METHOD Work : E_PROGRESS // commands TransportUnit to TRANSPORT_START
VAR_INPUT
  Execute     : BOOL;
END_VAR
VAR_INST
  _nErrorId   : UDINT;
  _eState     : E_PROGRESS;
END_VAR
//-----------------------------------------------------------------------------
IF NOT Execute 
THEN 
	_eState                       := E_PROGRESS.PROGRESS_INIT; 
END_IF 
//-----------------------------------------------------------------------------
IF NOT Check() 
THEN 
	Work                          := E_PROGRESS.PROGRESS_ERROR; 
	RETURN; 
END_IF
//-----------------------------------------------------------------------------
//-----------------------------------------------------------------------------
CASE _eState
OF
  E_PROGRESS.PROGRESS_INIT:
    IF Execute
    THEN
      _nErrorId                 := 0;

      _XtsTransportCtrl.Cmd     := E_XTS_TRANSPORT_CTRL.CMD_NULL;
      _eState                   := E_PROGRESS.PROGRESS_BUSY;

      IF (_MessageLevel > E_MessageType.eMessageError)
      THEN
        _stMsg.eType            := E_MessageType.eMessageInfo;
        _stMsg.eSubdevice       := e_Subdevice.Application_Work;
        _stMsg.iErrorNumber     := 0;
        _stMsg.sText            := concat(TO_STRING(_eState), ': ');
        f_MessageSet(_stMsg);
      END_IF
    END_IF
  //-----------------------------------------------------------------------------
  //-----------------------------------------------------------------------------
  E_PROGRESS.PROGRESS_BUSY:
    _XtsTransportCtrl.Cmd       := E_XTS_TRANSPORT_CTRL.CMD_TRANSPORT_START;

    IF (_XtsTransportState.State = E_XTS_TRANSPORT_STATE.TRANSPORT_START + E_PROGRESS.PROGRESS_ERROR)
    THEN
      _eState                   := E_PROGRESS.PROGRESS_ERROR;
      _nErrorId                 := _XtsTransportState.GroupInfo.GroupErrorId; 

    ELSIF (_XtsTransportState.State = E_XTS_TRANSPORT_STATE.TRANSPORT_START + E_PROGRESS.PROGRESS_DONE)
    THEN
      _eState                   := E_PROGRESS.PROGRESS_PREPARE;
    END_IF
  //-----------------------------------------------------------------------------
  // spare states: 
  //  - the work is done for the YardMaster
  //  - you can now work on the CTRL/STATE structures of the Instances
  //-----------------------------------------------------------------------------
  E_PROGRESS.PROGRESS_PREPARE:
    _eState                     := E_PROGRESS.PROGRESS_STARTUP;
  //---------------------------------------------------------------------------------------------------------------
  //---------------------------------------------------------------------------------------------------------------
  E_PROGRESS.PROGRESS_STARTUP:
    _eState                     := E_PROGRESS.PROGRESS_CHECK;
  //---------------------------------------------------------------------------------------------------------------
  //---------------------------------------------------------------------------------------------------------------
  E_PROGRESS.PROGRESS_CHECK:
    _eState                     := E_PROGRESS.PROGRESS_OCCUPIED;
  //---------------------------------------------------------------------------------------------------------------
  //---------------------------------------------------------------------------------------------------------------
  E_PROGRESS.PROGRESS_OCCUPIED:
    _eState                     := E_PROGRESS.PROGRESS_WORKING;
  //---------------------------------------------------------------------------------------------------------------
  //---------------------------------------------------------------------------------------------------------------
  E_PROGRESS.PROGRESS_WORKING:
    _eState                     := E_PROGRESS.PROGRESS_STILL_WORKING;
  //---------------------------------------------------------------------------------------------------------------
  //---------------------------------------------------------------------------------------------------------------
  E_PROGRESS.PROGRESS_STILL_WORKING:
    _eState                     := E_PROGRESS.PROGRESS_DONE;

    IF (_MessageLevel > E_MessageType.eMessageError)
    THEN
      _stMsg.eType              := E_MessageType.eMessageInfo;
      _stMsg.eSubdevice         := e_Subdevice.Application_Work;
      _stMsg.iErrorNumber       := 0;
      _stMsg.sText              := concat(TO_STRING(_eState), ': ');
      f_MessageSet(_stMsg);
    END_IF

END_CASE
//-----------------------------------------------------------------------------
//-----------------------------------------------------------------------------

Work                            := _eState;
END_METHOD

PROPERTY XtsTransportCtrl : REFERENCE TO ST_XTS_TRANSPORT_CTRL
SET
_XtsTransportCtrl REF= XtsTransportCtrl;
END_SET
END_PROPERTY

PROPERTY XtsTransportState : REFERENCE TO ST_XTS_TRANSPORT_STATE
SET
_XtsTransportState REF= XtsTransportState;
END_SET
END_PROPERTY

END_FUNCTION_BLOCK

// ---- _MSG/f_MessageSet.TcPOU
FUNCTION f_MessageSet : BOOL
VAR_INPUT
  stMessage     : ST_Message;
END_VAR
VAR
  _uiIndex      : UINT;
  _MainDevice   : e_Device;
  _nModRes      : UDINT;     // residual after modulo
END_VAR

stMessage.tTime                     := GVL_MSG_XTS.sLocalTime;

// why here? so all calls to this function may stay the same
_nModRes                            := stMessage.eDevice MOD e_Device.General;
_MainDevice                         := stMessage.eDevice - _nModRes;

CASE _MainDevice
OF
  //--------------------------------------------------------------------------------
  e_device.DataProduct:
    // this is your data, if you choose to use this message system
    FOR _uiIndex := 1 TO GVL_MSG_XTS.MAX_MESSAGE
    DO
      IF (GVL_MSG_XTS.ProductMessages[_uiIndex].eType = e_MessageType.eMessageEmpty)
      THEN
        GVL_MSG_XTS.ProductMessages[_uiIndex]      := stMessage;
        GVL_MSG_XTS.MessageProductIndex            := _uiIndex;
        EXIT;
      END_IF
    END_FOR
  
    IF (stMessage.eType = E_MessageType.eMessageError)
    THEN
      // in case of error: increment counter
      GVL_MSG_XTS.MessageProductError              := GVL_MSG_XTS.MessageProductError + 1;
    END_IF
  //--------------------------------------------------------------------------------
  e_Device.Process,
  e_Device.Application:
    FOR _uiIndex := 1 TO GVL_MSG_XTS.MAX_MESSAGE
    DO
      IF (GVL_MSG_XTS.ApplicationMessages[_uiIndex].eType = e_MessageType.eMessageEmpty)
      THEN
        GVL_MSG_XTS.ApplicationMessages[_uiIndex]  := stMessage;    // yes, we grab global values directly, only here
        GVL_MSG_XTS.MessageApplicationIndex        := _uiIndex;
        EXIT;
      END_IF
    END_FOR
    IF (stMessage.eType = E_MessageType.eMessageError)
    THEN
      // in case of error: increment counter
      GVL_MSG_XTS.MessageApplicationError          := GVL_MSG_XTS.MessageApplicationError + 1;
    END_IF
  //--------------------------------------------------------------------------------
  e_Device.MetricsXts:
    FOR _uiIndex := 1 TO GVL_MSG_XTS.MAX_MESSAGE
    DO
      IF (GVL_MSG_XTS.MetricsMessages[_uiIndex].eType = e_MessageType.eMessageEmpty)
      THEN
        GVL_MSG_XTS.MetricsMessages[_uiIndex]      := stMessage;    // yes, we grab global values directly, only here
        GVL_MSG_XTS.MessageMetricsIndex            := _uiIndex;
        EXIT;
      END_IF
    END_FOR
    IF (stMessage.eType = E_MessageType.eMessageError)
    THEN
      // in case of error: increment counter
      GVL_MSG_XTS.MessageMetricsError              := GVL_MSG_XTS.MessageMetricsError + 1;
    END_IF
  //--------------------------------------------------------------------------------
  e_Device.MetricsAxis:
    FOR _uiIndex := 1 TO GVL_MSG_XTS.MAX_MESSAGE
    DO
      IF (GVL_MSG_AXIS.MetricMessages[_uiIndex].eType = e_MessageType.eMessageEmpty)
      THEN
        GVL_MSG_AXIS.MetricMessages[_uiIndex]  := stMessage;    // yes, we grab global values directly, only here
        GVL_MSG_AXIS.MessageMetricIndex        := _uiIndex;
        EXIT;
      END_IF
    END_FOR
    IF (stMessage.eType = E_MessageType.eMessageError)
    THEN
      // in case of error: increment counter
      GVL_MSG_AXIS.MessageMetricError          := GVL_MSG_AXIS.MessageMetricError + 1;
    END_IF
  //--------------------------------------------------------------------------------
  e_Device.Axis,
  e_Device.XfcAxis,
  e_device.XfcTouchProbe,
  e_device.XfcTriggerBox,
  e_Device.Camming,
  e_device.NciChannel,
  e_device.NciChannelCtrl:
    FOR _uiIndex := 1 TO GVL_MSG_XTS.MAX_MESSAGE
    DO
      IF (GVL_MSG_AXIS.MotionMessages[_uiIndex].eType = e_MessageType.eMessageEmpty)
      THEN
        GVL_MSG_AXIS.MotionMessages[_uiIndex]  := stMessage;    // yes, we grab global values directly, only here
        GVL_MSG_AXIS.MessageMotionIndex        := _uiIndex;
        EXIT;
      END_IF
    END_FOR
    IF (stMessage.eType = E_MessageType.eMessageError)
    THEN
      // in case of error: increment counter
      GVL_MSG_AXIS.MessageMotionError           := GVL_MSG_AXIS.MessageMotionError + 1;
    END_IF
  //--------------------------------------------------------------------------------
ELSE
  CASE stMessage.eDevice
  OF
    Device_MainApplication,
    Device_XmlData,              
    Device_Utilities:
      FOR _uiIndex := 1 TO GVL_MSG_XTS.MAX_MESSAGE
      DO
        IF (GVL_MSG_XTS.ApplicationMessages[_uiIndex].eType = e_MessageType.eMessageEmpty)
        THEN
          GVL_MSG_XTS.ApplicationMessages[_uiIndex]:= stMessage;    // yes, we grab global values directly, only here
          GVL_MSG_XTS.MessageApplicationIndex      := _uiIndex;
          EXIT;
        END_IF
      END_FOR
      IF (stMessage.eType = E_MessageType.eMessageError)
      THEN
        // in case of error: increment counter
        GVL_MSG_XTS.MessageApplicationError        := GVL_MSG_XTS.MessageApplicationError + 1;
      END_IF

    Device_MainAxis,
    Device_Nci,
    Device_Cam,
    Device_Functions,
    Device_FlyingSaw,
    Device_ParameterSelector:     // PLC_MOTION
      FOR _uiIndex := 1 TO GVL_MSG_XTS.MAX_MESSAGE
      DO
        IF (GVL_MSG_AXIS.MotionMessages[_uiIndex].eType = e_MessageType.eMessageEmpty)
        THEN
          GVL_MSG_AXIS.MotionMessages[_uiIndex]:= stMessage;    // yes, we grab global values directly, only here
          GVL_MSG_AXIS.MessageMotionIndex      := _uiIndex;
          EXIT;
        END_IF
      END_FOR
      IF (stMessage.eType = E_MessageType.eMessageError)
      THEN
        // in case of error: increment counter
        GVL_MSG_AXIS.MessageMotionError        := GVL_MSG_AXIS.MessageMotionError + 1;
      END_IF

    Device_Main,
    Device_MoverSelector:
      FOR _uiIndex := 1 TO GVL_MSG_XTS.MAX_MESSAGE
      DO
        IF (GVL_MSG_XTS.TransportMessages[_uiIndex].eType = e_MessageType.eMessageEmpty)
        THEN
          GVL_MSG_XTS.TransportMessages[_uiIndex]  := stMessage;
          GVL_MSG_XTS.MessageTransportIndex        := _uiIndex;
          EXIT;
        END_IF
      END_FOR
  ELSE    
    //--------------------------------------------------------------------------------
    FOR _uiIndex := 1 TO GVL_MSG_XTS.MAX_MESSAGE
    DO
      IF (GVL_MSG_XTS.TransportMessages[_uiIndex].eType = e_MessageType.eMessageEmpty)
      THEN
        GVL_MSG_XTS.TransportMessages[_uiIndex]    := stMessage;
        GVL_MSG_XTS.MessageTransportIndex          := _uiIndex;
        EXIT;
      END_IF
    END_FOR
  
    IF (stMessage.eType = E_MessageType.eMessageError)
    THEN
      // in case of error: increment counter
      GVL_MSG_XTS.MessageTransportError := GVL_MSG_XTS.MessageTransportError + 1;
    END_IF
  END_CASE
END_CASE

END_FUNCTION

// ---- APPLICATION/_types/Instance/fb_Instance.TcPOU
//---------------------------------------------------------------------------------------------------------------
//
//  HAUD 2026.11.23
//
//
//---------------------------------------------------------------------------------------------------------------
//  fb_Instance
//---------------------------------------------------------------------------------------------------------------
//---------------------------------------------------------------------------------------------------------------
//  - base class for a process instance to work with fb_ProcessCollector
//  - extend this class to build top level transport logic
//    - example extension: fb_DistributorByTicket (1 to many)
//
//  What is it that I truly desire? 
//  --> to reduce the amount of handshakes that are required for a range of XtsStation
//  --> keep the granularity of a single station also for a range of stations
//  --> reuse existing interfaces
//
//  What an Instance is for:
//  - customized administrative transport related work
//    - reading of process tickets
//    - checking of queues
//    - handshaking ranges of stations
//      - automate handshake sequences with the collectors
//    - letting the stations write station tickets
//    - writing of process tickets
//
//  How an Instance is supposed to work:
//  - An Instance is of the same nature as a fb_StationProcess.Cycle / fb_ProcessCollector.Cycle
//    
//    --> you should build a Cycle() method
//    --> the default state after self init at PowerOn shall be a disabled state
//      --> a station behaviour follows the following concept:
//        - switch on --> station moves to enabled state
//        - enabled : switch to detection
//          - detection : detect what is given to you (e.g. QueueCount or LinkedList ticket)
//          - detected work leads to station asking for permission
//        - permitted : execute whatever is mandatory for starting the process (move to position etc)
//        - start / done
//          --> you decide how to handshake
//        - ready to send out : prepare your destination data here!
//        - send out : handshake sequence for safely permitting motion of a mover and transport of information
//
//    - It is up to you to decide how many handshakes with the CollectorInterface to automate in an instance
//      - example, a default distributor may require handshakes for every mover, 
//                 a mask driven distributor distributes until it has worked through the mask autonomously
//
//    - Read the existing extensions:
//      - you will find a 2-step progression for state changes
//      - they use the enumerations E_INSTANCE_CMD / E_INSTANCE_STATE
//        - in combination with E_PROGRESS
//        - there will be flowcharts for the existing extensions.
//
//---------------------------------------------------------------------------------------------------------------
//  - there are already 3 primitives available
//    - [1 to 1] DistributorByQueue
//      - a single station for 
//        - fly-by and change dynamics
//        - simple one stop
//
//    - [1 to m] DistributorByTicket
//      - a single station with ticket inbox check for
//        - sending a mover to a range of stations in accordance to the bitmask it received
//
//    - [m to 1] ProcessByTicket
//      - a range of stations handling a stationary process with ticket inbox
//      - single and nested stops
//      - sends movers to a single target (distributor)
//---------------------------------------------------------------------------------------------------------------
//
//---------------------------------------------------------------------------------------------------------------
//  - ProcessId : _nProcess --> whoami, this is me
//---------------------------------------------------------------------------------------------------------------
//
//  - who is required for my work on the outside?
//  - fb_ProcessCollector[_nProcess].Cycle() is called in MAIN_APP(PRG)
//    - provides interface
//    - handles range of XtsStations
//    - range must be closed and in consecutive order
//
//    - combines states into bitmasks, one bit per XtsStation
//    - controls forwarding of commands to range of XtsStations 
//      (see fb_ProcessCollector.Cycle())
//
//---------------------------------------------------------------------------------------------------------------
//  - CollectorInterface 
//---------------------------------------------------------------------------------------------------------------
//    - reference to all _ItfProcessCollector(I_ProcessCollector)[]
//    - _ItfProcessCollector[nProcess] carries ctrl/state information
//
//    - Control / State of the CollectorInterface
//      - local _stCollectorCtrl / _stCollectorState datafields are linked (REF=) to CollectorInterface.ProcessCtrl / .ProcessState
//        - since this connection shall be done automatically I put it in Check() method
//          --> see Check()
// 
//      - local datafield for control and state provided
//        - since CollectorInterface.ProcessCtrl and CollectorInterface.ProcessState are reference pointers
//          --> the real datafield has to come from somewhere, 
//              in this case the local datafields _stCollectorCtrl/_stCollectorState
//
//      - _stCollectorCtrl(ST_PROCESS_CTRL)
//        --> commands to the connected CollectorInterface;
//
//        Cmd               : E_PROCESS_CTRL; // command enum for collector
//        ProcessTarget     : UINT;           // target of my process
//        ActivateStation   : T_PROCESS;      // is checked for every job
//                                            // every bit is an XtsStation
//
//        NestMask          : BYTE;           // one mask for all XtsStations
//        - every bit is a PosStop within an XtsStation
//
//      - _stCollectorState(ST_PROCESS_STATE)
//        --> status information from the connected CollectorInterface
//        --> check for plausible StationLast / StationFirst range of XtsStations
//
//        State             : E_PROCESS_STATE;  // state enum from collector
//        Result            : E_PROGRESS;       // substate from collector, E_PROGRESS.PROGRESS_BUSY signals the collector state is ready for interaction
//                                              // fb_DistributorByTicket may give you an idea of the use of a substate 
//        Check             : E_PROCESS_CHECK;  // plausibility check of StationLast and StationFirst (the result of Check() --> _eCheck) 
//---------------------------------------------------------------------------------------------------------------
//  - InstanceCtrl(_stInstanceCtrl) 
//---------------------------------------------------------------------------------------------------------------
//  - incoming handshakes from higher up
//    - remember, 
//      this shall be a helper so you can do administrative stuff here 
//      so your actual process logic (picking, dispensing, syncing, gearing) may live elsewhere
// 
//---------------------------------------------------------------------------------------------------------------
//  - InstanceState(_stInstanceState)
//---------------------------------------------------------------------------------------------------------------
//  - reporting to higher up
//
//
//---------------------------------------------------------------------------------------------------------------
//---------------------------------------------------------------------------------------------------------------
//  - basic check and var names, so you can build your procedures with it
//
//  - processes may be connected via linked list, you decide.
//    - linked list for processes is intended to work as job buffer
//    - linked list provides information via ST_PROCESS_DATA, 
//      add what you have to in there
//    - linked list to all process instances provided
//
//  - inherit this base class for your application, call Check() every cycle at the top before you do anything
//       IF NOT Check() THEN 
//         RETURN; 
//       END_IF
//
//---------------------------------------------------------------------------------------------------------------//
// This SOFTWARE is provided as an Example by THE PROVIDER "as is" and "with all faults." THE PROVIDER makes no  //
// representations or warranties of any kind concerning the safety, suitability, lack of viruses, inaccuracies,  //
// typographical errors, or other harmful components of this SOFTWARE. There are inherent dangers in the use of  //
// any software, and you are solely responsible for determining whether this SOFTWARE is compatible with your    //
// equipment and other software installed on your equipment. You are also solely responsible for the protection  //
// of your equipment and backup of your data, and THE PROVIDER will not be liable for any damages you may suffer //
// in connection with using, modifying, or distributing this SOFTWARE.                                           //
//---------------------------------------------------------------------------------------------------------------//
FUNCTION_BLOCK ABSTRACT fb_Instance
VAR
  // process index
  _nProcess               : E_INSTANCE;           // whoami

  _stInstanceCtrl         : REFERENCE TO ARRAY[1..MAX_PROCESS] OF ST_INSTANCE_CTRL;
  _stInstanceState        : REFERENCE TO ARRAY[1..MAX_PROCESS] OF ST_INSTANCE_STATE;

  _eCmd,
  _eCmdOld                : E_INSTANCE_CMD;       // commands for local state machine
  _eStateInstance         : E_INSTANCE_STATE;     // local state machine for infeed procedure

  _eResult                : E_PROGRESS;           // result for methods
  _eStateProgress         : E_PROGRESS;           // substate for local state machine

  _eInit                  : E_PROGRESS;           // startup
  _eCheck                 : E_INSTANCE_CHECK;     // pointer checks

  // local ctrl / state datafields for you to use, connected by reference to _ItfProcessCollector[_nProcess]
  _stCollectorCtrl        : ST_PROCESS_CTRL;      // control to write, connected by reference to _ItfProcessCollector
  _stCollectorState       : ST_PROCESS_STATE;     // state   to read,  connected by reference to _ItfProcessCollector

  _ItfProcessCollector    : ARRAY[1..MAX_PROCESS] OF I_ProcessCollector;    // information and configuration of the connected ProcessCollector for given range of XtsStations

  _ItfProcessList         : ARRAY[1..MAX_PROCESS] OF I_Process_LinkedList;  // access to all linked lists for writing tickets
  _stListResult           : ST_PROCESS_LIST_RESULT;
  _stProcessData          : ST_PROCESS_DATA;

  {attribute 'displaymode':='bin'}
  _wTargetMask            : ARRAY[1..SIZEOF(T_PROCESS)*8] OF BYTE; // bits for PosStop[] to use in XtsStation of target process

  // position window within which a mover must be for the instance to react
  // value in abs modulo axis value
  //  - crossing the modulo turn is evaluated --> (Start > End) case is valid as window
  _rCheckPositionStart    : LREAL;
  _rCheckPositionEnd      : LREAL;

  _stMsg                  : ST_Message;
  _MessageLevel           : E_MessageType := E_MessageType.eMessageInfo;
END_VAR

METHOD Check : BOOL // call this method in the extending/inheriting class
//-----------------------------------------------------------------------------
//-----------------------------------------------------------------------------
// plausibility checks
//-----------------------------------------------------------------------------
IF NOT (_nProcess > 0)
THEN
  _eCheck                 := E_INSTANCE_CHECK.PROCESS_ID_ZERO;
  RETURN;
END_IF

IF NOT (_nProcess < E_INSTANCE.INSTANCE_MAX)
THEN
  _eCheck                 := E_INSTANCE_CHECK.PROCESS_ID_MAX;
  RETURN;
END_IF
//-----------------------------------------------------------------------------
//-----------------------------------------------------------------------------
// pointer checks
//-----------------------------------------------------------------------------
IF NOT __ISVALIDREF(_stInstanceCtrl)
THEN
  _eCheck                 := E_INSTANCE_CHECK.INVALID_INSTANCE_CONTROL_REFERENCE;
  RETURN;
END_IF

IF NOT __ISVALIDREF(_stInstanceState)
THEN
  _eCheck                 := E_INSTANCE_CHECK.INVALID_INSTANCE_STATE_REFERENCE;
  RETURN;
END_IF

IF NOT (_ItfProcessCollector[_nProcess] <> 0) 
THEN
  _eCheck                 := E_INSTANCE_CHECK.POINTER_COLLECTOR_ITF_INVALID;
  RETURN;
END_IF

IF NOT (_ItfProcessCollector[_nProcess].ProcessId > 0)
THEN
  _eCheck                 := E_INSTANCE_CHECK.PROCESS_ID_ZERO;
  RETURN;
END_IF

IF NOT (_ItfProcessCollector[_nProcess].ProcessId < E_INSTANCE.INSTANCE_MAX)
THEN
  _eCheck                 := E_INSTANCE_CHECK.PROCESS_ID_MAX;
  RETURN;
END_IF

IF NOT (_nProcess = _ItfProcessCollector[_nProcess].ProcessId)
THEN
  _eCheck                 := E_INSTANCE_CHECK.PROCESS_ID_NOTEQUAL_COLLECTOR_ID;
  RETURN;
END_IF

IF NOT (_ItfProcessList[_nProcess] <> 0)
THEN
  _eCheck                 := E_INSTANCE_CHECK.PROCESS_LIST_ITF_INDEX_INVALID;
  RETURN;
END_IF
//-----------------------------------------------------------------------------
//-----------------------------------------------------------------------------
// connect datafields to interface of ProcessCollector
//-----------------------------------------------------------------------------
_ItfProcessCollector[_nProcess].ProcessCtrl   REF= _stCollectorCtrl;
_ItfProcessCollector[_nProcess].ProcessState  REF= _stCollectorState;

//-----------------------------------------------------------------------------
//-----------------------------------------------------------------------------
// set message device
//-----------------------------------------------------------------------------
_stMsg.eDevice            := e_Device.Process + TO_UINT(_nProcess);
//-----------------------------------------------------------------------------
//-----------------------------------------------------------------------------
_eCheck                   := E_INSTANCE_CHECK.CHECK_DONE;
Check                     := TRUE;
END_METHOD

PROPERTY CheckPositionEnd : lreal // end of the position window to execute logic (should be higher than the WaitPos this instance is working on)
GET
CheckPositionEnd := _rCheckPositionEnd;
END_GET
SET
_rCheckPositionEnd := CheckPositionEnd;
END_SET
END_PROPERTY

PROPERTY CheckPositionStart : lreal // start of the position window to execute instance logic
GET
CheckPositionStart := _rCheckPositionStart;
END_GET
SET
_rCheckPositionStart := CheckPositionStart;
END_SET
END_PROPERTY

METHOD CmdLog

IF (_MessageLevel > E_MessageType.eMessageError)
THEN
  _stMsg.eSubdevice       := e_Subdevice.Instance_Command;
  _stMsg.iErrorNumber     := _nProcess;
  _stMsg.sText            := concat('E_INSTANCE_CMD', '.');
  _stMsg.sText            := concat(_stMsg.sText, TO_STRING(_eCmd));
  f_MessageSet(_stMsg);
END_IF
END_METHOD

PROPERTY CollectorInterface : array[1..MAX_PROCESS] of I_ProcessCollector
SET
_ItfProcessCollector := CollectorInterface;
END_SET
END_PROPERTY

PROPERTY InstanceCtrl : REFERENCE TO ARRAY[1..MAX_PROCESS] OF ST_INSTANCE_CTRL
SET
_stInstanceCtrl ref= InstanceCtrl;
END_SET
END_PROPERTY

PROPERTY InstanceState : REFERENCE TO ARRAY[1..MAX_PROCESS] OF ST_INSTANCE_STATE
SET
_stInstanceState ref= InstanceState;
END_SET
END_PROPERTY

PROPERTY MessageLevel : e_MessageType
GET
MessageLevel := _MessageLevel;
END_GET
SET
_MessageLevel := MessageLevel;

IF NOT (_eInit  = E_PROGRESS.PROGRESS_DONE) OR
   NOT (_eCheck = E_INSTANCE_CHECK.CHECK_DONE)
THEN
  RETURN;
ELSE
  _ItfProcessCollector[_nProcess].MessageLevel := _MessageLevel;
END_IF
END_SET
END_PROPERTY

PROPERTY ProcessId : E_INSTANCE
GET
ProcessId := _nProcess;
END_GET
SET
_nProcess := ProcessId;
END_SET
END_PROPERTY

PROPERTY ProcessLinkedLists : ARRAY[1..max_process] OF I_Process_LinkedList
SET
_ItfProcessList := ProcessLinkedLists;
END_SET
END_PROPERTY

END_FUNCTION_BLOCK

// ---- APPLICATION/Instances/fb_DistributorByQueue.TcPOU
//---------------------------------------------------------------------------------------------------------------
//
//  HAUD 2026.10.20
//
//
//  fb_DistributorByQueue
//  - uses 1 XtsStation via _ItfProcessCollector
//  - this instance only checks its queue after being enabled, then sends the mover to static station target (1 to 1)
//    - why only 1 to 1? 
//      --> this instance is intended to merely switch dynamics of a mover after the mover entered into the check window
//      --> change dynamics and off you go
//
//  - inherits fb_Instance, which provides a design pattern in order to build different specific processes in a structured way
//  - used for targeting movers to predetermined substation (one to one)
//  - the idea is to simply switch this instance off and on, the distributing is merely logic, 
//    so the handshakes are automated,
//      You enable first,
//      then acknowledge the outfeed 
//      and disable once the mover is dealt with (this part you might want to change if you do not need the feedback on the disabled state)
//      and back to enable to start all over again.
//
//
//  - constructed with fb_Instance main state (_eState) in addition to a substate (_eStateProgress)
//  - substate enables to handle procedures within main state by preventing race conditions 
//    with the help of small steps and decisions with clear separation from each other 
//
//---------------------------------------------------------------------------------------------------------------//
// This SOFTWARE is provided as an Example by THE PROVIDER "as is" and "with all faults." THE PROVIDER makes no  //
// representations or warranties of any kind concerning the safety, suitability, lack of viruses, inaccuracies,  //
// typographical errors, or other harmful components of this SOFTWARE. There are inherent dangers in the use of  //
// any software, and you are solely responsible for determining whether this SOFTWARE is compatible with your    //
// equipment and other software installed on your equipment. You are also solely responsible for the protection  //
// of your equipment and backup of your data, and THE PROVIDER will not be liable for any damages you may suffer //
// in connection with using, modifying, or distributing this SOFTWARE.                                           //
//---------------------------------------------------------------------------------------------------------------//
FUNCTION_BLOCK fb_DistributorByQueue EXTENDS fb_Instance
VAR
  _nProcessTarget               : E_INSTANCE;     // to whom am I connected

  // target XTS station range
  _nTargetStationLast           : UINT;           // where does the target process end
  _nTargetStationFirst          : UINT;           // where does the target process start

  _idx                          : UINT;
  _nTargetIndex                 : ARRAY[1..SIZEOF(T_PROCESS)*8] OF USINT; // helper var to copy to my process (_ItfProcessCollector[_nProcess].TargetIndex)

  _StationState                 : ST_STATION_STATE;   // A Distributor has only one XtsStation to work

  _nBatch                       : UDINT;
  _bUnmannedSender              : BOOL := TRUE;   // test var to test automated behaviour, so you only switch on/off
END_VAR

//-----------------------------------------------------------------------------
//-----------------------------------------------------------------------------
// check pointer and interface
// connect Ctrl/State to _ItfProcessCollector
// set message device identification
//-----------------------------------------------------------------------------
IF NOT Check() THEN 
  RETURN; 
END_IF
//-----------------------------------------------------------------------------
// check init command (hard reset)
//-----------------------------------------------------------------------------
_eCmd                                         := _stInstanceCtrl[_nProcess].Cmd;
IF (_eCmd <> _eCmdOld)
THEN
  CASE _eCmd
  OF
    E_INSTANCE_CMD.INIT:
      // clear init info
      _nBatch                                 := 0;
      _eInit                                  := _ItfProcessCollector[_nProcess].Init(FALSE);
  
      IF _ItfProcessList[_nProcess].InitList()  // clear linked list
      THEN
        Clear();
        _eStateInstance                       := E_INSTANCE_STATE.INIT;
        _eStateProgress                       := E_PROGRESS.PROGRESS_INIT;
      END_IF

    E_INSTANCE_CMD.CLEAR:
        _eStateInstance                       := E_INSTANCE_STATE.DISABLED;
        _eStateProgress                       := E_PROGRESS.PROGRESS_INIT;
  END_CASE
  CmdLog();
  _eCmdOld                                    := _eCmd;
END_IF
//-----------------------------------------------------------------------------
// cyclic information of station
//-----------------------------------------------------------------------------
_StationState                                 := _ItfProcessCollector[_nProcess].GetStationState  (_ItfProcessCollector[_nProcess].StationLast);
//-----------------------------------------------------------------------------
//-----------------------------------------------------------------------------
// state machine to send a mover as soon as added to the station's queue
//-----------------------------------------------------------------------------
CASE _eStateInstance // main state machine
OF
  E_INSTANCE_STATE.NULL:                      // first cycle init
    IF _ItfProcessList[_nProcess].InitList()
    THEN
      _eInit                                  := _ItfProcessCollector[_nProcess].Init(FALSE);
      _eStateProgress                         := E_PROGRESS.PROGRESS_INIT;
      _eStateInstance                         := E_INSTANCE_STATE.INIT;
    END_IF


  E_INSTANCE_STATE.INIT:                      // plausibility checks and _ItfProcessCollector Init
    //-------------------------------------------------------------------------
    CASE _eStateProgress
    OF
    //-------------------------------------------------------------------------
      E_PROGRESS.PROGRESS_ERROR:
        IF (_nProcessTarget > 0) AND
           (_nProcessTarget < E_INSTANCE.INSTANCE_MAX)
        THEN
          _eStateProgress                     := E_PROGRESS.PROGRESS_INIT;
        END_IF

    // E_INSTANCE_STATE.INIT:
    //-------------------------------------------------------------------------
      E_PROGRESS.PROGRESS_INIT:
        IF NOT (_nProcessTarget > 0) OR
           NOT (_nProcessTarget < E_INSTANCE.INSTANCE_MAX)
        THEN
          // an invalid target you must have not
          _eStateProgress                     := E_PROGRESS.PROGRESS_ERROR;
        ELSE
          _eStateProgress                     := E_PROGRESS.PROGRESS_BUSY;
        END_IF

    // E_INSTANCE_STATE.INIT:
    //-------------------------------------------------------------------------
      E_PROGRESS.PROGRESS_BUSY:
        // wait for my process collector check (_State.Check) to be done
        //  - checks range of XtsStations
        //  - checks count of XtsStations
        IF (_stCollectorState.Check = E_PROCESS_CHECK.CHECK_DONE)
        THEN
          _eInit                              := _ItfProcessCollector[_nProcess].Init(TRUE);
  
          IF (_eInit = E_PROGRESS.PROGRESS_DONE)
          THEN
            IF NOT (_nProcessTarget > 0) OR
               NOT (_nProcessTarget < E_INSTANCE.INSTANCE_MAX)
            THEN
              // an invalid target you must have not
              _eStateProgress                 := E_PROGRESS.PROGRESS_ERROR;

              _stMsg.eType                    := E_MessageType.eMessageError;
              _stMsg.eSubdevice               := e_Subdevice.Instance_DistributorByQueue;
              _stMsg.iErrorNumber             := _nProcessTarget;
              _stMsg.sText                    := concat(TO_STRING(_eStateInstance), ': ProcessTarget: ');
              _stMsg.sText                    := concat(_stMsg.sText, TO_STRING(_eStateProgress));
              f_MessageSet(_stMsg);

            ELSE
              _nTargetStationLast             := _ItfProcessCollector[_nProcessTarget].StationLast;
              _nTargetStationFirst            := _ItfProcessCollector[_nProcessTarget].StationFirst;

              // initialization of Infeed: _ItfProcessCollector with XtsStation
              _stCollectorCtrl.Cmd            := E_PROCESS_CTRL.PROCESS_DISABLE;  // first, switch off _ItfProcessCollector and XtsStation
              _eStateProgress                 := E_PROGRESS.PROGRESS_INIT;        // clear sub state
              _eStateInstance                 := E_INSTANCE_STATE.DISABLED;       // switch to disabled as default after startup
            END_IF
          END_IF
        END_IF
    END_CASE
END_CASE
//-----------------------------------------------------------------------------
//-----------------------------------------------------------------------------
// DISABLED:
//  - clear local list result data
//  - wait for enable from the outside
//  - wait for an entry in my list
//-----------------------------------------------------------------------------
CASE _eStateInstance
OF
  E_INSTANCE_STATE.DISABLED:
    //-------------------------------------------------------------------------
    CASE _eStateProgress
    OF
      E_PROGRESS.PROGRESS_INIT:
        _eStateProgress                       := E_PROGRESS.PROGRESS_BUSY;
        _stCollectorCtrl.ActivateStation      := 0;
        _stCollectorCtrl.NestMask             := 1;
        
    // E_INSTANCE_STATE.DISABLED:
    //-------------------------------------------------------------------------
      E_PROGRESS.PROGRESS_BUSY:
        //----------------------------------
        //  wait for command from higher up
        //----------------------------------
        CASE _eCmd
        OF
          E_INSTANCE_CMD.ENABLE:              // higher up decided to enable
            _eStateInstance                   := E_INSTANCE_STATE.DETECTION;
            _eStateProgress                   := E_PROGRESS.PROGRESS_BUSY;

  
            IF (_MessageLevel > E_MessageType.eMessageInfo)
            THEN
              _stMsg.eType                    := E_MessageType.eMessageVerbose;
              _stMsg.eSubdevice               := e_Subdevice.Instance_DistributorByQueue;
              _stMsg.iErrorNumber             := 0;
              _stMsg.sText                    := concat(TO_STRING(_eStateInstance), ': ');
              _stMsg.sText                    := concat(_stMsg.sText, TO_STRING(_eStateProgress));
              f_MessageSet(_stMsg);
            END_IF
        END_CASE
    END_CASE
END_CASE
//-----------------------------------------------------------------------------
// DETECTION: 
//  - check station queue
//  - switch on collector when mover is detected
//-----------------------------------------------------------------------------
CASE _eStateInstance
OF
  E_INSTANCE_STATE.DETECTION:
    //-------------------------------------------------------------------------
    CASE _eStateProgress
    OF
      E_PROGRESS.PROGRESS_BUSY:
        IF (_eCmd = E_INSTANCE_CMD.DISABLE)
        THEN
          _eStateInstance                     := E_INSTANCE_STATE.DISABLED;
          _eStateProgress                     := E_PROGRESS.PROGRESS_INIT;



        ELSIF (_StationState.nQueue > 0)
        THEN
          // as this instance is an automated sender to route movers, checking the queue is enough
          _eStateProgress                     := E_PROGRESS.PROGRESS_CHECK;

          IF (_MessageLevel > E_MessageType.eMessageError)
          THEN
            _stMsg.eType                      := E_MessageType.eMessageInfo;
            _stMsg.eSubdevice                 := e_Subdevice.Process_StationQueue_Check;
            _stMsg.iErrorNumber               := 0;
            _stMsg.sText                      := concat(TO_STRING(_eStateInstance), ': ');
            _stMsg.sText                      := concat(_stMsg.sText, '_StationState.nQueue: ');
            _stMsg.sText                      := concat(_stMsg.sText, TO_STRING(_StationState.nQueue));
            f_MessageSet(_stMsg);
          END_IF

          IF (_MessageLevel = E_MessageType.eMessageBatch)
          THEN
            _stMsg.eType                      := E_MessageType.eMessageBatch;
            _stMsg.eSubdevice                 := e_Subdevice.Instance_DistributorByQueue;
            _stMsg.iErrorNumber               := _StationState.nMoverId;
            _stMsg.sText                      := concat(TO_STRING(_eStateProgress), ': ');
            _stMsg.sText                      := concat(_stMsg.sText, TO_STRING(e_message_batch.MSG_BATCH_JOB_STARTED));
            f_MessageSet(_stMsg);
          END_IF
        END_IF
    END_CASE
    // E_INSTANCE_STATE.DETECTION
    //-------------------------------------------------------------------------
    CASE _eStateProgress
    OF
      E_PROGRESS.PROGRESS_CHECK:
        // check state of CollectorInterface
        CASE _stCollectorState.State
        OF
          E_PROCESS_STATE.PROCESS_DISABLE:

          CASE _stCollectorState.Result
          OF
            // busy from _State.Result means, waiting for input
            E_PROGRESS.PROGRESS_BUSY:
              // now the preparation for the target process may begin
              _stCollectorCtrl.Cmd               := E_PROCESS_CTRL.PROCESS_ENABLE;
              // I am a distributor (1 to 1), there is only one XtsStation to work
              _stCollectorCtrl.ActivateStation   := 1;

              _eStateInstance                 := E_INSTANCE_STATE.ENABLED;      // go check if my process is switched on
              _eStateProgress                 := E_PROGRESS.PROGRESS_INIT;      // reset substate

              IF (_MessageLevel > E_MessageType.eMessageInfo)
              THEN
                _stMsg.eType                  := E_MessageType.eMessageVerbose;
                _stMsg.eSubdevice             := e_Subdevice.Instance_DistributorByQueue;
                _stMsg.iErrorNumber           := 0;
                _stMsg.sText                  := concat(TO_STRING(_eStateInstance), ': ');
                _stMsg.sText                  := concat(_stMsg.sText, TO_STRING(_eStateProgress));
                f_MessageSet(_stMsg);
              END_IF
          END_CASE
        END_CASE
    END_CASE
END_CASE
//-----------------------------------------------------------------------------
// ENABLED
//  - check process for enabled station
//  - switch to infeed
//  - check if infeed is active
//  - allow movers to enter
//-----------------------------------------------------------------------------
CASE _eStateInstance
OF
  E_INSTANCE_STATE.ENABLED:
    //-------------------------------------------------------------------------
    CASE _eStateProgress
    OF
      E_PROGRESS.PROGRESS_INIT:
        CASE _stCollectorState.State
        OF
          E_PROCESS_STATE.PROCESS_ENABLE:
          CASE _stCollectorState.Result
          OF
            E_PROGRESS.PROGRESS_BUSY:
              // now my process and all XtsStations within are switched on
              // check infeed into my process
              _stCollectorCtrl.Cmd            := E_PROCESS_CTRL.PROCESS_STATIONS_INFEED; // tells my process to go check the infeed
              _eStateProgress                 := E_PROGRESS.PROGRESS_BUSY; // go check how the infeed into my process is doing

              IF (_MessageLevel > E_MessageType.eMessageInfo)
              THEN
                _stMsg.eType                  := E_MessageType.eMessageVerbose;
                _stMsg.eSubdevice             := e_Subdevice.Instance_DistributorByQueue;
                _stMsg.iErrorNumber           := 0;
                _stMsg.sText                  := concat(TO_STRING(_eStateInstance), ': ');
                _stMsg.sText                  := concat(_stMsg.sText, TO_STRING(_eStateProgress));
                f_MessageSet(_stMsg);
              END_IF
          END_CASE
        END_CASE
    END_CASE
    // E_INSTANCE_STATE.ENABLED:
    //-------------------------------------------------------------------------
    CASE _eStateProgress
    OF
      E_PROGRESS.PROGRESS_BUSY:
        CASE _stCollectorState.State
        OF
          E_PROCESS_STATE.PROCESS_STATIONS_INFEED:
          CASE _stCollectorState.Result
          OF
            E_PROGRESS.PROGRESS_BUSY:
              // now we know who wants to enter
              _stCollectorCtrl.Cmd            := E_PROCESS_CTRL.PROCESS_STATIONS_SEND;  // send mover to outfeed process
              _eStateProgress                 := E_PROGRESS.PROGRESS_PREPARE;           // go check sending of mover
  
              IF (_MessageLevel > E_MessageType.eMessageInfo)
              THEN
                _stMsg.eType                  := E_MessageType.eMessageVerbose;
                _stMsg.eSubdevice             := e_Subdevice.Instance_DistributorByQueue;
                _stMsg.iErrorNumber           := 0;
                _stMsg.sText                  := concat(TO_STRING(_eStateInstance), ': ');
                _stMsg.sText                  := concat(_stMsg.sText, TO_STRING(_eStateProgress));
                f_MessageSet(_stMsg);
              END_IF
          END_CASE
        END_CASE
    END_CASE
    // E_INSTANCE_STATE.ENABLED:
    //-------------------------------------------------------------------------
    CASE _eStateProgress
    OF
      E_PROGRESS.PROGRESS_PREPARE:
        CASE _stCollectorState.State
        OF
          E_PROCESS_STATE.PROCESS_STATIONS_OUTFEED:
          CASE _stCollectorState.Result
          OF
            E_PROGRESS.PROGRESS_BUSY:

              IF (_rCheckPositionEnd > _rCheckPositionStart)  // the default case
              THEN
                IF (_StationState.rMoverModPos > _rCheckPositionStart) AND
                   (_StationState.rMoverModPos < _rCheckPositionEnd)
                THEN
                  // mover is in range and can leave now
                  _eStateInstance             := E_INSTANCE_STATE.FINISH;     // go send mover
                  _eStateProgress             := E_PROGRESS.PROGRESS_INIT;    // reset substate
    
                  IF (_MessageLevel > E_MessageType.eMessageInfo)
                  THEN
                    _stMsg.eType              := E_MessageType.eMessageVerbose;
                    _stMsg.eSubdevice         := e_Subdevice.Instance_DistributorByQueue;
                    _stMsg.iErrorNumber       := _StationState.nMoverId;
                    _stMsg.sText              := concat(TO_STRING(_eStateInstance), ': D: ');
                    _stMsg.sText              := concat(_stMsg.sText, TO_STRING(_eStateProgress));
                    f_MessageSet(_stMsg);
                  END_IF
                END_IF
              ELSE
                // _rCheckPositionEnd < _rCheckPositionStart
                // the modulo turn crossing case
                IF (_StationState.rMoverModPos > _rCheckPositionStart) OR
                   (_StationState.rMoverModPos < _rCheckPositionEnd)
                THEN
                  // mover is in range and can leave now
                  _eStateInstance             := E_INSTANCE_STATE.FINISH;     // go send mover
                  _eStateProgress             := E_PROGRESS.PROGRESS_INIT;    // reset substate
    
                  IF (_MessageLevel > E_MessageType.eMessageInfo)
                  THEN
                    _stMsg.eType              := E_MessageType.eMessageVerbose;
                    _stMsg.eSubdevice         := e_Subdevice.Instance_DistributorByQueue;
                    _stMsg.iErrorNumber       := _StationState.nMoverId;
                    _stMsg.sText              := concat(TO_STRING(_eStateInstance), ': M: ');
                    _stMsg.sText              := concat(_stMsg.sText, TO_STRING(_eStateProgress));
                    f_MessageSet(_stMsg);
                  END_IF
                END_IF
              END_IF
          END_CASE
        END_CASE
    END_CASE
END_CASE
//-----------------------------------------------------------------------------
// FINISH:
//  - write target
//  - command outfeed of mover
//  - check disabled state of ControllerInterface proceed
//-----------------------------------------------------------------------------
CASE _eStateInstance
OF
  E_INSTANCE_STATE.FINISH:
    //-------------------------------------------------------------------------
    CASE _eStateProgress
    OF
      E_PROGRESS.PROGRESS_INIT:
        IF NOT _bUnmannedSender
        THEN
          _eStateProgress                     := E_PROGRESS.PROGRESS_BUSY;
        ELSE
          _eStateProgress                     := E_PROGRESS.PROGRESS_PREPARE;
        END_IF

        // the sending of mover
        _nTargetIndex[1]                      := TO_USINT(_nTargetStationLast);
        // write Xts target onto CollectorInterface
        _ItfProcessCollector[_nProcess].TargetIndex := _nTargetIndex;
  
        IF (_MessageLevel > E_MessageType.eMessageError)
        THEN
          _stMsg.eType                        := E_MessageType.eMessageInfo;
          _stMsg.eSubdevice                   := e_Subdevice.Instance_DistributorByQueue;
          _stMsg.iErrorNumber                 := _nTargetIndex[1];
          _stMsg.sText                        := concat('_nTargetIndex[1]: ', TO_STRING(_nTargetIndex[1]));
          _stMsg.sText                        := concat(_stMsg.sText, ' nMoverId: ');
          _stMsg.sText                        := concat(_stMsg.sText, TO_STRING(_StationState.nMoverId));
          f_MessageSet(_stMsg);
        END_IF
    END_CASE
    //-------------------------------------------------------------------------
    CASE _eStateProgress
    OF
      E_PROGRESS.PROGRESS_BUSY:
        CASE _stCollectorState.State
        OF
          // CollectorInterface is checking if mover is ready for outfeed
          E_PROCESS_STATE.PROCESS_STATIONS_OUTFEED:
          CASE _stCollectorState.Result
          OF
            // CollectorInterface gets busy when state of mover is confirmed
            // (_wStateOut = _wActivateStation)
            E_PROGRESS.PROGRESS_BUSY:
            // now data is prepared and copied to the right places

            //----------------------------------
            //  wait for command from higher up
            //----------------------------------
            CASE _eCmd
            OF
              E_INSTANCE_CMD.FINISH:          // send mover out!!
                _stCollectorCtrl.Cmd          := E_PROCESS_CTRL.PROCESS_STATIONS_OUTFEED; // release the kraken!
                _eStateProgress               := E_PROGRESS.PROGRESS_DONE;                // mover is on its way

                IF (_MessageLevel = E_MessageType.eMessageBatch)
                THEN
                  _stMsg.eType                := E_MessageType.eMessageBatch;
                  _stMsg.eSubdevice           := e_Subdevice.Instance_DistributorByQueue;
                  _stMsg.iErrorNumber         := _StationState.nMoverId;
                  _stMsg.sText                := concat(TO_STRING(_eStateProgress), ': ');
                  _stMsg.sText                := concat(_stMsg.sText, TO_STRING(e_message_batch.MSG_BATCH_JOB_DONE));
                  f_MessageSet(_stMsg);
                END_IF

                // increment internal debug counter 
                _nBatch                       := _nBatch + 1;
            END_CASE
          END_CASE
        END_CASE
    END_CASE
    //-------------------------------------------------------------------------
    CASE _eStateProgress
    OF
      E_PROGRESS.PROGRESS_PREPARE:
        CASE _stCollectorState.State
        OF
          // CollectorInterface is checking if mover is ready for outfeed
          E_PROCESS_STATE.PROCESS_STATIONS_OUTFEED:
            CASE _stCollectorState.Result
            OF
              // CollectorInterface gets busy when state of mover is confirmed
              // (_wStateOut = _wActivateStation)
              E_PROGRESS.PROGRESS_BUSY:
              // now data is prepared and copied to the right places
                _stCollectorCtrl.Cmd          := E_PROCESS_CTRL.PROCESS_STATIONS_OUTFEED; // release the kraken!
                _eStateProgress               := E_PROGRESS.PROGRESS_CHECK;                // mover is on its way
  
                IF (_MessageLevel = E_MessageType.eMessageBatch)
                THEN
                  _stMsg.eType                := E_MessageType.eMessageBatch;
                  _stMsg.eSubdevice           := e_Subdevice.Instance_DistributorByQueue;
                  _stMsg.iErrorNumber         := _StationState.nMoverId;
                  _stMsg.sText                := concat(TO_STRING(_eStateProgress), ': ');
                  _stMsg.sText                := concat(_stMsg.sText, TO_STRING(e_message_batch.MSG_BATCH_JOB_DONE));
                  f_MessageSet(_stMsg);
                END_IF
                  // increment internal debug counter 
                _nBatch                       := _nBatch + 1;
            END_CASE
        END_CASE
    END_CASE
    //-------------------------------------------------------------------------
    CASE _eStateProgress
    OF
      E_PROGRESS.PROGRESS_CHECK:
        CASE _stCollectorState.State
        OF
          // the last command has released the mover,
          // CollectorInterface checks:
          //  - if the mover has left the station (_wStateOut = 0)
          //  --> return to disabled state.
          E_PROCESS_STATE.PROCESS_DISABLE:
            CASE _stCollectorState.Result
            OF
              // CollectorInterface is disabled and has no mover in control
              E_PROGRESS.PROGRESS_BUSY:
                _eStateInstance               := E_INSTANCE_STATE.DISABLED;
                _eStateProgress               := E_PROGRESS.PROGRESS_INIT;
  
                IF (_MessageLevel > E_MessageType.eMessageError)
                THEN
                  _stMsg.eType                := E_MessageType.eMessageInfo;
                  _stMsg.eSubdevice           := e_Subdevice.Instance_DistributorByQueue;
                  _stMsg.iErrorNumber         := 1;
                  _stMsg.sText                := TO_STRING(_eStateInstance);
                  _stMsg.sText                := concat(_stMsg.sText, ': ');
                  _stMsg.sText                := concat(_stMsg.sText, TO_STRING(_eStateProgress));
                  f_MessageSet(_stMsg);
                END_IF
            END_CASE
        END_CASE
    END_CASE
    //-------------------------------------------------------------------------
    CASE _eStateProgress
    OF
      E_PROGRESS.PROGRESS_DONE:
        CASE _stCollectorState.State
        OF
          // the last command has released the mover,
          // CollectorInterface checks:
          //  - if the mover has left the station (_wStateOut = 0)
          //  --> return to disabled state.
          E_PROCESS_STATE.PROCESS_DISABLE:
          CASE _stCollectorState.Result
          OF
            // CollectorInterface is disabled and has no mover in control
            E_PROGRESS.PROGRESS_BUSY:
              //----------------------------------
              //  wait for command from higher up
              //----------------------------------
              CASE _eCmd
              OF
                // your command to disable is required
                E_INSTANCE_CMD.DISABLE:
                  _eStateInstance             := E_INSTANCE_STATE.DISABLED;
                  _eStateProgress             := E_PROGRESS.PROGRESS_INIT;

                  IF (_MessageLevel > E_MessageType.eMessageError)
                  THEN
                    _stMsg.eType              := E_MessageType.eMessageInfo;
                    _stMsg.eSubdevice         := e_Subdevice.Instance_DistributorByQueue;
                    _stMsg.iErrorNumber       := 0;
                    _stMsg.sText              := TO_STRING(_eStateInstance);
                    _stMsg.sText              := concat(_stMsg.sText, ': ');
                    _stMsg.sText              := concat(_stMsg.sText, TO_STRING(_eStateProgress));
                    f_MessageSet(_stMsg);
                  END_IF

              END_CASE
          END_CASE
        END_CASE
    END_CASE
    //-------------------------------------------------------------------------
END_CASE
//-----------------------------------------------------------------------------
//-----------------------------------------------------------------------------
_stInstanceState[_nProcess].ProcessIdentity   := _nProcess;
_stInstanceState[_nProcess].ProcessState      := _eStateInstance;
_stInstanceState[_nProcess].ProcessProgress   := _eStateProgress;
//-----------------------------------------------------------------------------
//-----------------------------------------------------------------------------
_stInstanceState[_nProcess].CollectorState    := _stCollectorState.State;
_stInstanceState[_nProcess].CollectorProgress := _stCollectorState.Result;
_stInstanceState[_nProcess].CollectorCheck    := _stCollectorState.Check;
_stInstanceState[_nProcess].StationCount      := _ItfProcessCollector[_nProcess].StationCount;
_stInstanceState[_nProcess].QueueProcessCount := _ItfProcessCollector[_nProcess].QueueProcessCount;
_stInstanceState[_nProcess].ListCount         := TO_UINT(_ItfProcessList[_nProcess].Count);
//-----------------------------------------------------------------------------
//-----------------------------------------------------------------------------

METHOD Clear : BOOL
VAR_INPUT
END_VAR
memset(ADR(_nTargetIndex), 0, SIZEOF(_nTargetIndex));

//_eStateInstance                         := E_INSTANCE_STATE.DISABLED;
_eStateProgress                 := E_PROGRESS.PROGRESS_INIT;

Clear                           := TRUE;
END_METHOD

PROPERTY ProcessTarget : E_INSTANCE
GET
ProcessTarget := _nProcessTarget;
END_GET
SET
_nProcessTarget := ProcessTarget;
END_SET
END_PROPERTY

END_FUNCTION_BLOCK

// ---- APPLICATION/Instances/fb_DistributorByTicket.TcPOU
//---------------------------------------------------------------------------------------------------------------
//
//  HAUD 2026.10.20
//
//
//  fb_DistributorByTicket
//  - uses 1 XtsStation via _ItfProcessCollector
//  - this instance checks its process list for an entry (Count > 0)
//      - pops ticket data from top of the list (GetHead)
//      - sends the mover to target stations according to bitmask in ST_PROCESS_DATA.wTarget
//
//  - inherits fb_Instance, which provides a design pattern in order to build different specific processes in a structured way
//  - used for targeting movers to predetermined bitmask of substations (one to many)
//
//
//  - constructed with fb_Instance main state (_eState) in addition to a substate (_eStateProgress)
//  - substate enables to handle procedures within main state by preventing race conditions 
//    with the help of small steps and decisions with clear separation from each other 
//
//---------------------------------------------------------------------------------------------------------------//
// This SOFTWARE is provided as an Exemple by THE PROVIDER "as is" and "with all faults." THE PROVIDER makes no  //
// representations or warranties of any kind concerning the safety, suitability, lack of viruses, inaccuracies,  //
// typographical errors, or other harmful components of this SOFTWARE. There are inherent dangers in the use of  //
// any software, and you are solely responsible for determining whether this SOFTWARE is compatible with your    //
// equipment and other software installed on your equipment. You are also solely responsible for the protection  //
// of your equipment and backup of your data, and THE PROVIDER will not be liable for any damages you may suffer //
// in connection with using, modifying, or distributing this SOFTWARE.                                           //
//---------------------------------------------------------------------------------------------------------------//
FUNCTION_BLOCK fb_DistributorByTicket EXTENDS fb_Instance
VAR
  //----------------------------------------------------------------------------------
  // outfeed target must be initialized with a valid target
  // I just use the default target that I am going to use in the basic process setup
  // this target is then updated and checked on arrival of a process ticket
  //----------------------------------------------------------------------------------
  _nProcessTarget               : E_INSTANCE;     // to whom am I connected --> to the data from the ticket
  //----------------------------------------------------------------------------------

  // target XTS station range
  _nTargetStationLast           : UINT;           // where does the target process end
  _nTargetStationFirst          : UINT;           // where does the target process start

  _WriteResult                  : ST_PROCESS_LIST_RESULT;   // last job written to target
  _DeleteResult                 : ST_PROCESS_LIST_RESULT;   // last job executed

  _nPrc                         : E_INSTANCE;
  _nTarget                      : E_INSTANCE;

  _idx                          : UINT;
  _nTargetIndex                 : ARRAY[1..SIZEOF(T_PROCESS)*8] OF USINT;

  _MoverInfo                    : ST_MOVER_INFO;      // Information from the Mover in Station
  _StationState                 : ST_STATION_STATE;   // BufferInfeed has only one XtsStation to work
END_VAR

//-----------------------------------------------------------------------------
//-----------------------------------------------------------------------------
// check pointer and interface
// connect Ctrl/State to _ItfProcessCollector
// set message device identification
//-----------------------------------------------------------------------------
IF NOT Check() THEN 
  RETURN; 
END_IF
//-----------------------------------------------------------------------------
// check command
//-----------------------------------------------------------------------------
_eCmd                                         := _stInstanceCtrl[_nProcess].Cmd;
IF (_eCmd <> _eCmdOld)
THEN
  CASE _eCmd
  OF
    E_INSTANCE_CMD.INIT:
      // clear init info
      _eInit                                  := _ItfProcessCollector[_nProcess].Init(FALSE);
  
      IF _ItfProcessList[_nProcess].InitList()  // clear linked list
      THEN
        Clear();
        _eStateInstance                       := E_INSTANCE_STATE.INIT;
        _eStateProgress                       := E_PROGRESS.PROGRESS_INIT;
      END_IF
  END_CASE
  CmdLog();
  _eCmdOld                                    := _eCmd;
END_IF
//-----------------------------------------------------------------------------
// cyclic information of mover and station
//-----------------------------------------------------------------------------
_StationState                                 := _ItfProcessCollector[_nProcess].GetStationState  (_ItfProcessCollector[_nProcess].StationLast);
//-----------------------------------------------------------------------------
//-----------------------------------------------------------------------------
// state machine for BufferInfeed work
//-----------------------------------------------------------------------------
CASE _eStateInstance
OF
  E_INSTANCE_STATE.NULL:
    // first cycle startup
    // initialize linked list, clears all entries
    IF _ItfProcessList[_nProcess].InitList()
    THEN
      _eInit                                  := _ItfProcessCollector[_nProcess].Init(FALSE);
      _eStateProgress                         := E_PROGRESS.PROGRESS_INIT;
      _eStateInstance                         := E_INSTANCE_STATE.INIT;
    END_IF


  E_INSTANCE_STATE.INIT:
    //-------------------------------------------------------------------------
    CASE _eStateProgress
    OF
    // E_INSTANCE_STATE.INIT:
    //-------------------------------------------------------------------------
      E_PROGRESS.PROGRESS_ERROR:
        IF (_nProcessTarget > 0) AND
           (_nProcessTarget < E_INSTANCE.INSTANCE_MAX)
        THEN
          _eStateProgress                     := E_PROGRESS.PROGRESS_INIT;
        END_IF

    // E_INSTANCE_STATE.INIT:
    //-------------------------------------------------------------------------
      E_PROGRESS.PROGRESS_INIT:
        IF NOT (_nProcessTarget > 0) OR
           NOT (_nProcessTarget < E_INSTANCE.INSTANCE_MAX)
        THEN
          _eStateProgress                     := E_PROGRESS.PROGRESS_ERROR;

        ELSE
          _eStateProgress                     := E_PROGRESS.PROGRESS_BUSY;
        END_IF

    // E_INSTANCE_STATE.INIT:
    //-------------------------------------------------------------------------
      E_PROGRESS.PROGRESS_BUSY:
        // wait for process collector check to be done
        //  - checks range of XtsStations
        //  - checks count of XtsStations
        IF (_stCollectorState.Check = E_PROCESS_CHECK.CHECK_DONE)
        THEN
          _eInit                              := _ItfProcessCollector[_nProcess].Init(TRUE);
  
          IF (_eInit = E_PROGRESS.PROGRESS_DONE)
          THEN
            IF NOT (_nProcessTarget > 0) OR
               NOT (_nProcessTarget < E_INSTANCE.INSTANCE_MAX)
            THEN
              // an invalid target you must have not
              _eStateProgress                 := E_PROGRESS.PROGRESS_ERROR;

              _stMsg.eType                    := E_MessageType.eMessageError;
              _stMsg.eSubdevice               := e_Subdevice.Instance_DistributorByTicket;
              _stMsg.iErrorNumber             := _nProcessTarget;
              _stMsg.sText                    := concat(TO_STRING(_eStateInstance), ': ProcessTarget: ');
              _stMsg.sText                    := concat(_stMsg.sText, TO_STRING(_eStateProgress));
              f_MessageSet(_stMsg);

            ELSE
              _ItfProcessCollector[_nProcess].Init(FALSE); // clear init procedure

              // initialization of BufferInfeed: _ItfProcessCollector with XtsStation
              _stCollectorCtrl.Cmd            := E_PROCESS_CTRL.PROCESS_DISABLE;  // switch off _ItfProcessCollector and XtsStation
              _eStateProgress                 := E_PROGRESS.PROGRESS_INIT;        // clear sub state
              _eStateInstance                 := E_INSTANCE_STATE.DISABLED;       // switch to disabled as default after startup
            END_IF
          END_IF
        END_IF
    END_CASE
END_CASE
//-----------------------------------------------------------------------------
// DISABLED:
//  - clear local list result data
//  - wait for enable from the outside
//-----------------------------------------------------------------------------
CASE _eStateInstance
OF
  E_INSTANCE_STATE.DISABLED:
    //-------------------------------------------------------------------------
    CASE _eStateProgress
    OF
      E_PROGRESS.PROGRESS_INIT:
        _stCollectorCtrl.Cmd                  := E_PROCESS_CTRL.PROCESS_DISABLE;  // switch off _ItfProcessCollector and XtsStation
        _eStateProgress                       := E_PROGRESS.PROGRESS_BUSY;
        // clear data for a new round
        memset(ADR(_stListResult), 0, SIZEOF(_stListResult));

        _stCollectorCtrl.ActivateStation      := 0; // clear activation mask of my process
        _stCollectorCtrl.NestMask             := 1; // my process target has one nest

        _nPrc                                 := _nProcess;
        _nTarget                              := _nProcessTarget;
    END_CASE
    // E_INSTANCE_STATE.DISABLED:
    //-------------------------------------------------------------------------
    CASE _eStateProgress
    OF
      E_PROGRESS.PROGRESS_BUSY:
        CASE _eCmd
        OF
          E_INSTANCE_CMD.ENABLE:              // turn it on!!
            _nPrc                             := _nProcess;
            _nTarget                          := _nProcessTarget;

            _eStateInstance                   := E_INSTANCE_STATE.DETECTION;
            _eStateProgress                   := E_PROGRESS.PROGRESS_BUSY;
  
            IF (_MessageLevel > E_MessageType.eMessageInfo)
            THEN
              _stMsg.eType                    := E_MessageType.eMessageVerbose;
              _stMsg.eSubdevice               := e_Subdevice.Instance_DistributorByTicket;
              _stMsg.iErrorNumber             := 0;
              _stMsg.sText                    := concat(TO_STRING(_eStateInstance), ': ');
              _stMsg.sText                    := concat(_stMsg.sText, TO_STRING(_eStateProgress));
              f_MessageSet(_stMsg);
            END_IF

        END_CASE
    END_CASE
END_CASE
//-----------------------------------------------------------------------------
// DETECTION: 
//  - check inked list and GetHead()
//  - copy job data
//  - switch on process
//-----------------------------------------------------------------------------
CASE _eStateInstance
OF
  E_INSTANCE_STATE.DETECTION:
    //-------------------------------------------------------------------------
    CASE _eStateProgress
    OF
      E_PROGRESS.PROGRESS_BUSY:
        IF (_eCmd = E_INSTANCE_CMD.DISABLE)
        THEN
          _eStateInstance                     := E_INSTANCE_STATE.DISABLED;
          _eStateProgress                     := E_PROGRESS.PROGRESS_INIT;

        ELSIF (_ItfProcessList[_nPrc].Count > 0)
        THEN
          // get new job order for my process
          // check my list for a new round of movers
          _stListResult                       := _ItfProcessList[_nPrc].GetHead();  // the list results carries information about the requirements of the target process (who and where)

          IF (_stListResult.wState <> 0)
          THEN
            // error in list results must not appear
            // if you land here, there is somethng wrong with the initialization or configuration of the linked list
            _eStateProgress                   := E_PROGRESS.PROGRESS_ERROR;

            _stMsg.eType                      := E_MessageType.eMessageError;
            _stMsg.eSubdevice                 := e_Subdevice.Process_LinkedList_GetHead;
            _stMsg.iErrorNumber               := _stListResult.wState;
            _stMsg.sText                      := concat(TO_STRING(_eStateInstance), ': _ListResult.wState: ');
            _stMsg.sText                      := concat(_stMsg.sText, TO_STRING(_eStateProgress));
            f_MessageSet(_stMsg);

          ELSE
            IF (_MessageLevel > E_MessageType.eMessageError)
            THEN
              _stMsg.eType                    := E_MessageType.eMessageInfo;
              _stMsg.eSubdevice               := e_Subdevice.Process_LinkedList_GetHead;
              _stMsg.iErrorNumber             := _nPrc;
              _stMsg.sText                    := concat(TO_STRING(_eStateInstance), ': ');
              _stMsg.sText                    := concat(_stMsg.sText, '_ListResult.stData.wTarget: ');
              _stMsg.sText                    := concat(_stMsg.sText, _ItfProcessCollector[_nPrc].BitsToString(_stListResult.stData.wTarget));
              f_MessageSet(_stMsg);
            END_IF

            _stProcessData                    := _stListResult.stData;  // list result contains data for target process

            IF (_stProcessData.wTarget > 0)
            THEN
              _eStateProgress                 := E_PROGRESS.PROGRESS_CHECK;

              IF (_MessageLevel = E_MessageType.eMessageBatch)
              THEN
                _stMsg.eType                  := E_MessageType.eMessageBatch;
                _stMsg.eSubdevice             := e_Subdevice.Instance_DistributorByTicket;
                _stMsg.iErrorNumber           := _nPrc;
                _stMsg.sText                  := concat(TO_STRING(_eStateProgress), ': ');
                _stMsg.sText                  := concat(_stMsg.sText, TO_STRING(e_message_batch.MSG_BATCH_JOB_STARTED));
                f_MessageSet(_stMsg);
              END_IF
            ELSE
              _DeleteResult                   := _ItfProcessList[_nPrc].RemoveHeadValue();
            END_IF

            // check target mask for entries
            IF NOT (_stProcessData.wTarget > 0)
            THEN
              _stMsg.eType                    := E_MessageType.eMessageWarning;
              _stMsg.eSubdevice               := e_Subdevice.Instance_DistributorByTicket;
              _stMsg.iErrorNumber             := 666;
              _stMsg.sText                    := concat(TO_STRING(_eStateInstance), ': ');
              _stMsg.sText                    := concat(_stMsg.sText, '_ProcessData.wTarget: ');
              _stMsg.sText                    := concat(_stMsg.sText, _ItfProcessCollector[_nProcess].BitsToString(_stProcessData.wTarget));
              f_MessageSet(_stMsg);
            END_IF
          END_IF
        END_IF
    END_CASE
    // E_INSTANCE_STATE.DETECTION
    //-------------------------------------------------------------------------
    CASE _eStateProgress
    OF
      E_PROGRESS.PROGRESS_CHECK:
        // do some plausibility checks on the ticket data
        IF NOT (_stProcessData.nTargetId > 0) OR
           NOT (_stProcessData.nTargetId < E_INSTANCE.INSTANCE_MAX) OR
           NOT (_stProcessData.nTargetId <> _nProcess)
        THEN
          _stMsg.eType                        := E_MessageType.eMessageError;
          _stMsg.eSubdevice                   := e_Subdevice.Instance_DistributorByTicket;
          _stMsg.iErrorNumber                 := _stProcessData.nTargetId;
          _stMsg.sText                        := concat(TO_STRING(_eStateInstance), ': _stProcessData.nTargetId: ');
          _stMsg.sText                        := concat(_stMsg.sText, TO_STRING(E_PROGRESS.PROGRESS_ERROR));
          f_MessageSet(_stMsg);

          // not a plausible target, delete ticket and go back to checking the list
          _DeleteResult                       := _ItfProcessList[_nPrc].RemoveHeadValue();
          _eStateProgress                     := E_PROGRESS.PROGRESS_BUSY;
        ELSE
          // update target data with ticket data
          _nTarget                            := _stProcessData.nTargetId;
          _nTargetStationLast                 := _ItfProcessCollector[_nTarget].StationLast;
          _nTargetStationFirst                := _ItfProcessCollector[_nTarget].StationFirst;

          IF (_ItfProcessCollector[_nTarget].ProcessState.Check = E_PROCESS_CHECK.CHECK_DONE)
          THEN
            _eStateProgress                   := E_PROGRESS.PROGRESS_WORKING;

            IF (_MessageLevel > E_MessageType.eMessageWarning)
            THEN
              _stMsg.eType                    := E_MessageType.eMessageInfo;
              _stMsg.eSubdevice               := e_Subdevice.Instance_DistributorByTicket;
              _stMsg.iErrorNumber             := _stProcessData.nTargetId;
              _stMsg.sText                    := concat(TO_STRING(_stProcessData.nProcessId), ': _stProcessData.nTargetId: ');
              _stMsg.sText                    := concat(_stMsg.sText, TO_STRING(_stProcessData.nTargetId));
              f_MessageSet(_stMsg);
            END_IF
          END_IF
        END_IF
    END_CASE
    // E_INSTANCE_STATE.DETECTION
    //-------------------------------------------------------------------------
    CASE _eStateProgress
    OF
      E_PROGRESS.PROGRESS_WORKING:
        // check for disabled process interface state
        CASE _stCollectorState.State
        OF
          E_PROCESS_STATE.PROCESS_DISABLE:

          CASE _stCollectorState.Result
          OF
            E_PROGRESS.PROGRESS_BUSY:         // busy from _State.Result means, waiting for input
              // now the preparation for the target process may begin
              _stCollectorCtrl.Cmd               := E_PROCESS_CTRL.PROCESS_ENABLE; // switch on my state machine in _ItfProcessCollector
              _stCollectorCtrl.ActivateStation   := 1;                             // enable my XtsStation in _ItfProcessCollector (BufferInfeed has only one XtsStation)

              _eStateInstance                 := E_INSTANCE_STATE.ENABLED;         // go check if my process is switched on
              _eStateProgress                 := E_PROGRESS.PROGRESS_INIT;         // reset substate

              IF (_MessageLevel > E_MessageType.eMessageInfo)
              THEN
                _stMsg.eType                  := E_MessageType.eMessageVerbose;
                _stMsg.eSubdevice             := e_Subdevice.Instance_DistributorByTicket;
                _stMsg.iErrorNumber           := 0;
                _stMsg.sText                  := concat(TO_STRING(_eStateInstance), ': ');
                _stMsg.sText                  := concat(_stMsg.sText, TO_STRING(_eStateProgress));
                f_MessageSet(_stMsg);
              END_IF
          END_CASE
        END_CASE
    END_CASE
END_CASE
//-----------------------------------------------------------------------------
// ENABLED
//  - check process for enabled stations from list entry
//  - switch to sending
//  - allow movers to be sent
//-----------------------------------------------------------------------------
CASE _eStateInstance
OF
  E_INSTANCE_STATE.ENABLED:
    //-------------------------------------------------------------------------
    CASE _eStateProgress
    OF
      E_PROGRESS.PROGRESS_INIT:
        CASE _stCollectorState.State
        OF
          E_PROCESS_STATE.PROCESS_ENABLE:
          CASE _stCollectorState.Result
          OF
            E_PROGRESS.PROGRESS_BUSY:
              // now my process and all XtsStations within are switched on
              // check infeed into my process
              _stCollectorCtrl.Cmd            := E_PROCESS_CTRL.PROCESS_STATIONS_SEND; // tells my process to go check the infeed
              _eStateProgress                 := E_PROGRESS.PROGRESS_BUSY; // go check how the infeed into my process is doing

              IF (_MessageLevel > E_MessageType.eMessageInfo)
              THEN
                _stMsg.eType                  := E_MessageType.eMessageVerbose;
                _stMsg.eSubdevice             := e_Subdevice.Instance_DistributorByTicket;
                _stMsg.iErrorNumber           := _StationState.nMoverId;
                _stMsg.sText                  := concat(TO_STRING(_eStateInstance), ': _stCollectorCtrl.Cmd: ');
                _stMsg.sText                  := concat(_stMsg.sText, TO_STRING(_stCollectorCtrl.Cmd));
                f_MessageSet(_stMsg);
              END_IF
          END_CASE
        END_CASE
    END_CASE
    // E_INSTANCE_STATE.ENABLED:
    //-------------------------------------------------------------------------
    CASE _eStateProgress
    OF
      E_PROGRESS.PROGRESS_BUSY:
        CASE _stCollectorState.State
        OF
          E_PROCESS_STATE.PROCESS_STATIONS_OUTFEED:
          CASE _stCollectorState.Result       // if collector is ready to send mover
          OF
            E_PROGRESS.PROGRESS_BUSY:
              // check if the mover is in range
              IF (_rCheckPositionEnd > _rCheckPositionStart)
              THEN
                IF (_StationState.rMoverModPos > _rCheckPositionStart) AND
                   (_StationState.rMoverModPos < _rCheckPositionEnd)
                THEN
                  _eStateProgress             := E_PROGRESS.PROGRESS_PREPARE;
                END_IF
              ELSE
                IF (_StationState.rMoverModPos > _rCheckPositionStart) OR
                   (_StationState.rMoverModPos < _rCheckPositionEnd)
                THEN
                  _eStateProgress             := E_PROGRESS.PROGRESS_PREPARE;
                END_IF
              END_IF
          END_CASE
        END_CASE
    END_CASE
    // E_INSTANCE_STATE.ENABLED:
    //-------------------------------------------------------------------------
    CASE _eStateProgress
    OF
      E_PROGRESS.PROGRESS_PREPARE:
        // now we know the mover is in range
        // continue to finish
        _stCollectorCtrl.Cmd                  := E_PROCESS_CTRL.PROCESS_STATIONS_SEND;

        _eStateInstance                       := E_INSTANCE_STATE.FINISH;   // go get data ready for outfeed
        _eStateProgress                       := E_PROGRESS.PROGRESS_INIT;  // reset substate
    END_CASE
END_CASE
//-----------------------------------------------------------------------------
// FINISH:
//  - write target (Last to First)
//  - delete target bit from linked list result (_ProcessData.wTarget)
//  - send out mover
//  - check _ProcessData.wTarget for next mover
//  - check if all movers in job were sent (ProcessData.wTarget = 0)
//  - RemoveHead() from my list
//  - AddTail() at TargetProcess
//  - check to proceed
//-----------------------------------------------------------------------------
CASE _eStateInstance
OF
  E_INSTANCE_STATE.FINISH:
    //-------------------------------------------------------------------------
    CASE _eStateProgress
    OF
      E_PROGRESS.PROGRESS_INIT:
      // check bit mask for sending mover to required targets
      // get target index for mover from process list entry
      FOR _idx := _nTargetStationLast TO _nTargetStationFirst BY(-1)
      DO
        IF (ItfProcessCollector[_nPrc].BitGet(_stProcessData.wTarget, _idx-_nTargetStationFirst))
        THEN
          _eStateProgress                     := E_PROGRESS.PROGRESS_BUSY;

          _nTargetIndex[1]                    := TO_USINT(_idx);
          _ItfProcessCollector[_nPrc].TargetIndex := _nTargetIndex; // write Xts target onto my ProcessCollector interface

          // got the target, now delete the just found bit of this job
          _stProcessData.wTarget              := _ItfProcessCollector[_nPrc].
                                                 BitDel(_stProcessData.wTarget, _idx-_nTargetStationFirst);

          IF (_MessageLevel > E_MessageType.eMessageInfo)
          THEN
            _stMsg.eType                      := E_MessageType.eMessageVerbose;
            _stMsg.eSubdevice                 := e_Subdevice.Instance_DistributorByTicket;
            _stMsg.iErrorNumber               := _idx;
            _stMsg.sText                      := concat('_ProcessData.wTarget: ', 
                                                 _ItfProcessCollector[_nPrc].BitsToString(_stProcessData.wTarget));
            f_MessageSet(_stMsg);
          END_IF
          IF (_MessageLevel > E_MessageType.eMessageError)
          THEN
            _stMsg.eType                        := E_MessageType.eMessageInfo;
            _stMsg.eSubdevice                   := e_Subdevice.Instance_DistributorByTicket;
            _stMsg.iErrorNumber                 := _StationState.nMoverId;
            _stMsg.sText                        := concat(TO_STRING(_eStateInstance), ': _nTargetIndex[1]: ');
            _stMsg.sText                        := concat(_stMsg.sText, TO_STRING(_idx));
            f_MessageSet(_stMsg);
          END_IF
          EXIT;
        END_IF
      END_FOR
    END_CASE
    // E_INSTANCE_STATE.FINISH:
    //-------------------------------------------------------------------------
    CASE _eStateProgress
    OF
      E_PROGRESS.PROGRESS_BUSY:
        CASE _stCollectorState.State
        OF
          E_PROCESS_STATE.PROCESS_STATIONS_OUTFEED: // double check my process' state
          CASE _stCollectorState.Result
          OF
            E_PROGRESS.PROGRESS_BUSY:
              // now data is prepared and copied to the right places
              _stCollectorCtrl.Cmd            := E_PROCESS_CTRL.PROCESS_STATIONS_OUTFEED; // tell my process to release the mover
              _eStateProgress                 := E_PROGRESS.PROGRESS_CHECK; // go check for more to do

              IF (_MessageLevel > E_MessageType.eMessageInfo)
              THEN
                _stMsg.eType                  := E_MessageType.eMessageVerbose;
                _stMsg.eSubdevice             := e_Subdevice.Instance_DistributorByTicket;
                _stMsg.iErrorNumber           := _nPrc;
                _stMsg.sText                  := concat(TO_STRING(_eStateInstance), ': ');
                _stMsg.sText                  := concat(_stMsg.sText, TO_STRING(_eStateProgress));
                f_MessageSet(_stMsg);
              END_IF
          END_CASE
        END_CASE
    END_CASE
    // E_INSTANCE_STATE.FINISH:
    //-------------------------------------------------------------------------
    CASE _eStateProgress
    OF
      E_PROGRESS.PROGRESS_CHECK:
        CASE _stCollectorState.State
        OF
          E_PROCESS_STATE.PROCESS_DISABLE:
            IF (_stProcessData.wTarget <> 0)
            THEN
              _stCollectorCtrl.Cmd               := E_PROCESS_CTRL.PROCESS_ENABLE; // switch on my state machine in _ItfProcessCollector
              _stCollectorCtrl.ActivateStation   := 1;                             // enable my XtsStation in _ItfProcessCollector (BufferInfeed has only one XtsStation)

              _eStateInstance                 := E_INSTANCE_STATE.ENABLED;         // go check if my process is switched on
              _eStateProgress                 := E_PROGRESS.PROGRESS_INIT;         // reset substate

              IF (_MessageLevel > E_MessageType.eMessageInfo)
              THEN
                _stMsg.eType                  := E_MessageType.eMessageVerbose;
                _stMsg.eSubdevice             := e_Subdevice.Instance_DistributorByTicket;
                _stMsg.iErrorNumber           := _nPrc;
                _stMsg.sText                  := concat(TO_STRING(_eStateInstance), ': ');
                _stMsg.sText                  := concat(_stMsg.sText, TO_STRING(_eStateProgress));
                f_MessageSet(_stMsg);
              END_IF
            ELSE
              // job done, all movers were sent
              // job done, delete from top of my list
              _DeleteResult                   := _ItfProcessList[_nPrc].RemoveHeadValue();

              IF (_DeleteResult.wState <> 0)
              THEN
                // deleting from list must be successful
                // IF you land here, there is something wrong with initialization or configuration of the linked list
                _eStateProgress               := E_PROGRESS.PROGRESS_ERROR;
              ELSE
                _eStateProgress               := E_PROGRESS.PROGRESS_WORKING; // job is done, now go and write ticket to _nTargetProcess

                IF (_MessageLevel > E_MessageType.eMessageError)
                THEN
                  _stMsg.eType                := E_MessageType.eMessageInfo;
                  _stMsg.eSubdevice           := e_Subdevice.Process_LinkedList_RemoveHead;
                  _stMsg.iErrorNumber         := 0;
                  _stMsg.sText                := concat(TO_STRING(_eStateInstance), ': ');
                  _stMsg.sText                := concat(_stMsg.sText, TO_STRING(_eStateProgress));
                  f_MessageSet(_stMsg);
                END_IF
              END_IF
            END_IF 
        END_CASE
    END_CASE
    // E_INSTANCE_STATE.FINISH:
    //-------------------------------------------------------------------------
    CASE _eStateProgress
    OF
      E_PROGRESS.PROGRESS_WORKING:
        // write process ticket, then go back up
        //_WriteResult                          := _ItfProcessList[_nTarget].AddTailValue(_stListResult.stData);

        IF (_WriteResult.wState <> 0)
        THEN
          // adding to target list must be successful on the first try
          // IF you land here, there is something wrong with initialization or configuration of the linked list
          _eStateProgress                     := E_PROGRESS.PROGRESS_ERROR;
        ELSE
          _eStateProgress                     := E_PROGRESS.PROGRESS_DONE;

          IF (_MessageLevel > E_MessageType.eMessageError)
          THEN
            _stMsg.eType                      := E_MessageType.eMessageInfo;
            _stMsg.eSubdevice                 := e_Subdevice.Process_LinkedList_AddTail;
            _stMsg.iErrorNumber               := _nTarget;
            _stMsg.sText                      := concat(TO_STRING(_eStateInstance), ': ');
            _stMsg.sText                      := concat(_stMsg.sText, TO_STRING(_eStateProgress));
            //f_MessageSet(_stMsg);
          END_IF
          IF (_MessageLevel = E_MessageType.eMessageBatch)
          THEN
            _stMsg.eType                      := E_MessageType.eMessageBatch;
            _stMsg.eSubdevice                 := e_Subdevice.Instance_DistributorByTicket;
            _stMsg.iErrorNumber               := _nPrc;
            _stMsg.sText                      := concat(TO_STRING(_eStateProgress), ': ');
            _stMsg.sText                      := concat(_stMsg.sText, TO_STRING(e_message_batch.MSG_BATCH_JOB_DONE));
            f_MessageSet(_stMsg);
          END_IF
        END_IF
    END_CASE
    // E_INSTANCE_STATE.FINISH:
    //-------------------------------------------------------------------------
    CASE _eStateProgress
    OF
      E_PROGRESS.PROGRESS_DONE:
        //----------------------------------
        //  wait for command from higher up
        //----------------------------------
        CASE _eCmd
        OF
          // command to disable required
          E_INSTANCE_CMD.DISABLE:
            _eStateInstance                   := E_INSTANCE_STATE.DISABLED;
            _eStateProgress                   := E_PROGRESS.PROGRESS_INIT;

            IF (_MessageLevel > E_MessageType.eMessageInfo)
            THEN
              _stMsg.eType                    := E_MessageType.eMessageVerbose;
              _stMsg.eSubdevice               := e_Subdevice.Instance_DistributorByTicket;
              _stMsg.iErrorNumber             := _nPrc;
              _stMsg.sText                    := concat(TO_STRING(_eStateInstance), ': ');
              _stMsg.sText                    := concat(_stMsg.sText, TO_STRING(_eStateProgress));
              f_MessageSet(_stMsg);
            END_IF
        END_CASE
    END_CASE
END_CASE
//-----------------------------------------------------------------------------
//-----------------------------------------------------------------------------
_stInstanceState[_nProcess].ProcessIdentity   := _nProcess;
_stInstanceState[_nProcess].ProcessState      := _eStateInstance;
_stInstanceState[_nProcess].ProcessProgress   := _eStateProgress;
//-----------------------------------------------------------------------------
//-----------------------------------------------------------------------------
_stInstanceState[_nProcess].CollectorState    := _stCollectorState.State;
_stInstanceState[_nProcess].CollectorProgress := _stCollectorState.Result;
_stInstanceState[_nProcess].CollectorCheck    := _stCollectorState.Check;
_stInstanceState[_nProcess].StationCount      := _ItfProcessCollector[_nProcess].StationCount;
_stInstanceState[_nProcess].QueueProcessCount := _ItfProcessCollector[_nProcess].QueueProcessCount;
_stInstanceState[_nProcess].ListCount         := TO_UINT(_ItfProcessList[_nProcess].Count);
//-----------------------------------------------------------------------------
//-----------------------------------------------------------------------------

METHOD Clear : BOOL
VAR_INPUT
END_VAR
memset(ADR(_nTargetIndex), 0, SIZEOF(_nTargetIndex));

//_eStateInstance                         := E_INSTANCE_STATE.DISABLED;
_eStateProgress                 := E_PROGRESS.PROGRESS_INIT;

Clear                           := TRUE;
END_METHOD

PROPERTY ProcessTarget : E_INSTANCE
GET
ProcessTarget := _nProcessTarget;
END_GET
SET
_nProcessTarget := ProcessTarget;
END_SET
END_PROPERTY

END_FUNCTION_BLOCK

// ---- APPLICATION/Instances/fb_ProcessByTicket.TcPOU
//---------------------------------------------------------------------------------------------------------------
//
//  HAUD 2026.10.25
//
//
//  fb_ProcessByTicket
//  - inherits fb_Instance
//
//  - uses range XtsStations via _ItfProcessCollector
//    - commands infeed of movers into stations for processing
//    - mask for stations asking for entry is double checked with mask in process ticket
//    - the sequence: 
//        enable [enables and detects work], 
//        work   [allows infeed and waits for all movers to arrive], 
//        finish [sends out movers writes outfeed ticket and disables]
//
//  - used for targeting movers to one predetermined target (many to one)
//    - the incoming ticket sets the target 
//      --> _nTargetOutfeed  := _stProcessData.nTargetId
//
//    - this instance can write a copy of the process ticket to an upstream DistributorByTicket
//      - write ticket to distributor on infeed  before process (optional if e_instance > 0)
//
//  - what about sending the ticket downstream?
//    - the target of this class is always a single station
//      --> DistributorByQueue does not need a ticket
//      --> DistributorByTicket is getting its ticket
//          a - from the Conductor via the extern ticket list
//          b - from a process downstram that knows how many and where the movers must be placed next
//
//  - processes are connected via linked list
//    - entry in list is detected
//    - entry in list determines count and place of used XtsStations in target process
//
//
//  - constructed with fb_Instance main state (_eState) in addition to a substate (_eStateProgress)
//  - substate enables to handle procedures within main state by preventing race conditions 
//    with the help of small steps and decisions with clear separation from each other 
//
//---------------------------------------------------------------------------------------------------------------//
// This SOFTWARE is provided as an Example by THE PROVIDER "as is" and "with all faults." THE PROVIDER makes no  //
// representations or warranties of any kind concerning the safety, suitability, lack of viruses, inaccuracies,  //
// typographical errors, or other harmful components of this SOFTWARE. There are inherent dangers in the use of  //
// any software, and you are solely responsible for determining whether this SOFTWARE is compatible with your    //
// equipment and other software installed on your equipment. You are also solely responsible for the protection  //
// of your equipment and backup of your data, and THE PROVIDER will not be liable for any damages you may suffer //
// in connection with using, modifying, or distributing this SOFTWARE.                                           //
//---------------------------------------------------------------------------------------------------------------//
FUNCTION_BLOCK fb_ProcessByTicket EXTENDS fb_Instance
VAR
  //----------------------------------------------------------------------------------
  // INFEED TARGET:  MAY BE UPDATED/CHANGED BEFORE SWITCHING TO E_INSTANCE_CMD.ENABLE
  //----------------------------------------------------------------------------------
  //  - sending a copy of the incoming ticket is done/tested
  //     the moment the ticket is detected
  //
  //    --> to be sent or not to be sent
  //        - that is best answered during E_INSTANCE_STATE.DISABLED
  //
  //  - (_nProcessTargetInfeed = INSTANCE_NULL) --> targeting deactivated
  //----------------------------------------------------------------------------------
  _nProcessTargetInfeed         : E_INSTANCE;     // to whom am I connected before work (set property for that)

  //----------------------------------------------------------------------------------
  // OUTFEED TARGET: must be initialized with a valid target
  //----------------------------------------------------------------------------------
  // The intent to have one valid setting for initialization, 
  //  the ticket data is checked on arrival and has dedicated messages in place
  // I just use the default target that I am going to use in the basic process setup
  //  - see MAIN_APP.eInit state machine as example
  //
  // OUTFEED TARGET: is updated and checked on arrival of a process ticket
  //----------------------------------------------------------------------------------
  _nProcessTargetOutfeed        : E_INSTANCE;     // to whom am I connected after  work --> to the data from the ticket
  //----------------------------------------------------------------------------------

  // target XTS station range
  _nTargetStationLast           : UINT;           // where does the target process end
  _nTargetStationFirst          : UINT;           // where does the target process start

  _WriteResult                  : ST_PROCESS_LIST_RESULT;   // last job written to target
  _DeleteResult                 : ST_PROCESS_LIST_RESULT;   // last job executed

  _idx                          : UINT;
  _nPrc                         : E_INSTANCE;
  _nTargetInfeed,
  _nTargetOutfeed               : E_INSTANCE;
  _nTargetIndex                 : ARRAY[1..SIZEOF(T_PROCESS)*8] OF USINT; // helper var to copy to my process (_ItfProcessCollector[_nProcess].TargetIndex)
  _StationState                 : ST_STATION_STATE;
END_VAR

//-----------------------------------------------------------------------------
//-----------------------------------------------------------------------------
// check pointer and interface
// connect Ctrl/State to _ItfProcessCollector
// set message device identification
//-----------------------------------------------------------------------------
IF NOT Check() THEN 
  RETURN; 
END_IF
//-----------------------------------------------------------------------------
// check init command (hard reset)
//-----------------------------------------------------------------------------
_eCmd                                         := _stInstanceCtrl[_nProcess].Cmd;
IF (_eCmd <> _eCmdOld)
THEN
  CASE _eCmd
  OF
    E_INSTANCE_CMD.INIT:
      // clear init info
      _eInit                                  := _ItfProcessCollector[_nProcess].Init(FALSE);
  
      IF _ItfProcessList[_nProcess].InitList()  // clear linked list
      THEN
        Clear();
        _eStateInstance                       := E_INSTANCE_STATE.INIT;
        _eStateProgress                       := E_PROGRESS.PROGRESS_INIT;
      END_IF
  END_CASE
  CmdLog();
  _eCmdOld                                    := _eCmd;
END_IF
//-----------------------------------------------------------------------------
// cyclic information of mover and station
//-----------------------------------------------------------------------------
_StationState                                 := _ItfProcessCollector[_nProcess].GetStationState  (_ItfProcessCollector[_nProcess].StationFirst);
//-----------------------------------------------------------------------------
// state machine for Infeed functionality
//-----------------------------------------------------------------------------
CASE _eStateInstance // main state machine
OF
  E_INSTANCE_STATE.NULL:                      // first cycle init
    IF _ItfProcessList[_nProcess].InitList()
    THEN
      _eInit                                  := _ItfProcessCollector[_nProcess].Init(FALSE);
      _eStateProgress                         := E_PROGRESS.PROGRESS_INIT;
      _eStateInstance                         := E_INSTANCE_STATE.INIT;
    END_IF


  E_INSTANCE_STATE.INIT:                      // plausibility checks and _ItfProcessCollector Init
    //-------------------------------------------------------------------------
    CASE _eStateProgress
    OF
    // E_INSTANCE_STATE.INIT:
    //-------------------------------------------------------------------------
      E_PROGRESS.PROGRESS_INIT:
        IF NOT (_nProcessTargetOutfeed > 0) OR
           NOT (_nProcessTargetOutfeed < E_INSTANCE.INSTANCE_MAX)
        THEN
          // an invalid target you must have not
          _eStateProgress                     := E_PROGRESS.PROGRESS_ERROR;
        ELSE
          _eStateProgress                     := E_PROGRESS.PROGRESS_BUSY;
        END_IF

